(* IEC 61131-3 sources: codesys-framework/txt/application/WeVe Core (library)/20 Service/I_Service, 2 files *)

(* ---- Initialize.method.st ---- *)
// Eenmalig bij de opstart. TRUE = klaar.
METHOD Initialize : BOOL
VAR_INPUT
END_VAR

(* ---- Reset.method.st ---- *)
// TRUE = reset gelukt.
METHOD Reset : BOOL
VAR_INPUT
END_VAR
